// TIA Portal V20 export
Screen "Pop-up_PRODDATA_PC_LEGEND_Popup"  330x409
  ScreenItem "Background" at 0,0 size 330x409  Type=HmiRectangle
  ScreenItem "Textfeld_Legende" at 1,1 size 328x25  Type=HmiTextBox
  ScreenItem "Cancel Mode" at 239,1 size 90x60  Type=HmiButton
  ScreenItem "Textfeld_11" at 65,308 size 260x96  Type=HmiTextBox
  ScreenItem "Textfeld_8" at 10,362 size 55x30  Type=HmiTextBox
  ScreenItem "Textfeld_9" at 23,343 size 30x20  Type=HmiTextBox
  ScreenItem "Textfeld_13" at 10,314 size 55x30  Type=HmiTextBox
  ScreenItem "Textfeld_10" at 10,34 size 208x28  Type=HmiTextBox
  ScreenItem "Textfeld_12" at 10,100 size 208x25  Type=HmiTextBox
  ScreenItem "Textfeld_14" at 10,63 size 315x35  Type=HmiTextBox
  ScreenItem "Textfeld_15" at 10,126 size 315x40  Type=HmiTextBox
  ScreenItem "Textfeld_2" at 10,168 size 55x30  Type=HmiTextBox
  ScreenItem "Textfeld_3" at 70,168 size 255x70  Type=HmiTextBox
  ScreenItem "Textfeld_4" at 10,201 size 55x30  Type=HmiTextBox
  ScreenItem "Textfeld_5" at 10,241 size 55x30  Type=HmiTextBox
  ScreenItem "Textfeld_6" at 70,238 size 255x70  Type=HmiTextBox
  ScreenItem "Textfeld_7" at 10,274 size 55x30  Type=HmiTextBox
